{attribute 'qualified_only'}
VAR_GLOBAL
	command : HmiCommand;
	status : HmiStatus;
END_VAR

(* stored: Version 1.1.0.1, ProductVersion 3.1.4026.12
   GVL RobotHmi: Id {b5fc5b2e-5306-5327-be70-30e2b1f2d258} *)
